Fanuc KAREL source: kx00004.KL

PROGRAM KX00004
%STACKSIZE=65535
%PRIORITY=65535
%NOLOCKGROUP
VAR
I : INTEGER
J : INTEGER
B : BOOLEAN
F : FILE
S : STRING[80]
P : XYZWPR
BEGIN
-- UNRESOLVED_PC line 11 opcodes [22 3F 3F 3D] marker_code=0
-- UNRESOLVED_PC line 12 opcodes [22 22 9C 9C 38 2C] marker_code=31
CLOSE FILE F
END KX00004
